// TIA Portal V20 export
DATA_BLOCK "01_Alle_Zaehler_DB"   // DB162
// stored: AssignedProDiagFB Pos12_ProDiag, InstanceOfName 01_Alle_Zaehler, InstanceOfType FB
"01_Alle_Zaehler"
   // VAR
   //    Zaehlsignal_Gesamt : Bool;
   //    Zaehlsignal_IO : Bool;
   //    Zaehlsignal_NIO : Bool;
   //    Zaehlsignal_NIO_LabView : Bool;
   //    "Zaehlsignal_IO_1 Palette 1" : Bool;
   //    "Zaehlsignal_IO_2 Palette 2" : Bool;
   //    "Zaehlsignal_IO_3 Palette 3" : Bool;
   //    "Zaehlsignal_IO_4 Palette 4" : Bool;
   //    "Zaehlsignal_IO_5 Palette 5" : Bool;
   //    "Zaehlsignal_NIO_1_Palette NIO" : Bool;
   //    Zaehlsignal_NIO_2 : Bool;
   //    Zaehlsignal_NIO_3 : Bool;
   //    Zaehlsignal_NIO_4 : Bool;
   //    Zaehlsignal_NIO_5 : Bool;
   //    Zaehlsignal_NIO_6 : Bool;
   // END_VAR
BEGIN
END_DATA_BLOCK
